(* PLC project case, CODESYS CODESYS V3.5 SP17 Patch 3 *)
(* stored: creationDateTime 2026-10-20T00:00:00 *)

CONFIGURATION Device
  RESOURCE Application ON PLC
    TASK MainTask(INTERVAL := T#20ms, PRIORITY := 5);
    TASK SlowTask(INTERVAL := T#20ms, PRIORITY := 10);
    PROGRAM PRG_A WITH MainTask : PRG_A;
    PROGRAM PRG_A WITH SlowTask : PRG_A;
  END_RESOURCE
END_CONFIGURATION
